FUNCTION_BLOCK EL_Template (* TEMPLATE for the rules of your equipment, EL_<Equipment>: copy it under that name, then change what says YOUR OWN, and this comment; keep the rest as it is. The logic of an equipment block: one holder at a time, outputs switched off before new ones go on, all off on release or abort, inputs reported when they change. Technical: Template: output values from its holder -> outputs (break before make); one holder at a time; all off on release or when the module aborts; inputs -> state channel when they change *)
  (* Standard: 61499-2 *)
  (* Version 0.1, 2026-09-28, Project contributors, AAU Smart Production Lab *)
  PACKAGE stoppering;
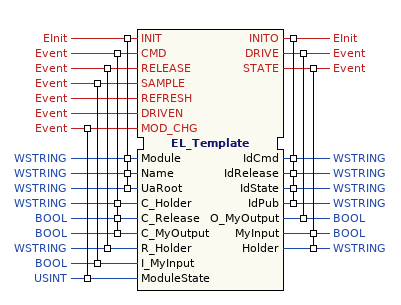
  EVENT_INPUT
    INIT : EInit WITH Module, Name, UaRoot; (* Initialise, once at start-up (the INIT chain); takes the values given with it *)
    CMD WITH C_Holder, C_Release, C_MyOutput; (* A command arrived from a holder *)
    RELEASE WITH R_Holder; (* A release arrived on the module's release channel (R_Holder) *)
    SAMPLE WITH I_MyInput; (* The inputs were read *)
    REFRESH; (* Cycle: write the outputs again *)
    DRIVEN; (* The outputs were written *)
    MOD_CHG WITH ModuleState; (* The module's state changed (its Aborting switches all off) *)
  END_EVENT
  EVENT_OUTPUT
    INITO : EInit WITH IdCmd, IdRelease, IdState, IdPub; (* Initialised: the next block of the INIT chain goes on *)
    DRIVE WITH O_MyOutput; (* Write the outputs *)
    STATE WITH MyInput, Holder; (* Publish the state (the inputs and the holder) *)
  END_EVENT
  VAR_INPUT
    Module : WSTRING; (* The module's name; its local channels are named after it (loc[<Module>/...]) *)
    Name : WSTRING; (* The equipment item's name: its local channels and OPC UA folder *)
    UaRoot : WSTRING; (* The module's OPC UA folder, e.g. /Objects/Filling *)
    C_Holder : WSTRING; (* Who sends the command *)
    C_Release : BOOL; (* Give up the equipment after this command *)
    C_MyOutput : BOOL; (* YOUR OWN, one per output pin. Commanded value of MyOutput *)
    R_Holder : WSTRING; (* Who gives up the equipment *)
    I_MyInput : BOOL; (* YOUR OWN, one per input pin. MyInput as read or received *)
    ModuleState : USINT; (* PackML state: 1 Clearing, 2 Stopped, 3 Starting, 4 Idle, 6 Execute, 7 Stopping, 8 Aborting, 9 Aborted, 15 Resetting *)
  END_VAR
  VAR_OUTPUT
    IdCmd : WSTRING; (* Local channel of the commands *)
    IdRelease : WSTRING; (* Local channel of the releases (the module's, one for all equipment) *)
    IdState : WSTRING; (* Local channel of the state *)
    IdPub : WSTRING; (* OPC UA ID of the published inputs *)
    O_MyOutput : BOOL; (* YOUR OWN, one per output pin. The value to write to MyOutput *)
    MyInput : BOOL; (* YOUR OWN, one per input pin. Template: MyInput, an input *)
    Holder : WSTRING; (* Who holds the equipment (empty: free) *)
  END_VAR
  VAR
    Publish : BOOL;
    Beat : USINT;
    LastHolder : WSTRING;
    Pending : BOOL;
    OffPending : BOOL;
    L_MyInput : BOOL; (* YOUR OWN, one per input pin *)
    N_MyOutput : BOOL; (* YOUR OWN, one per output pin *)
  END_VAR
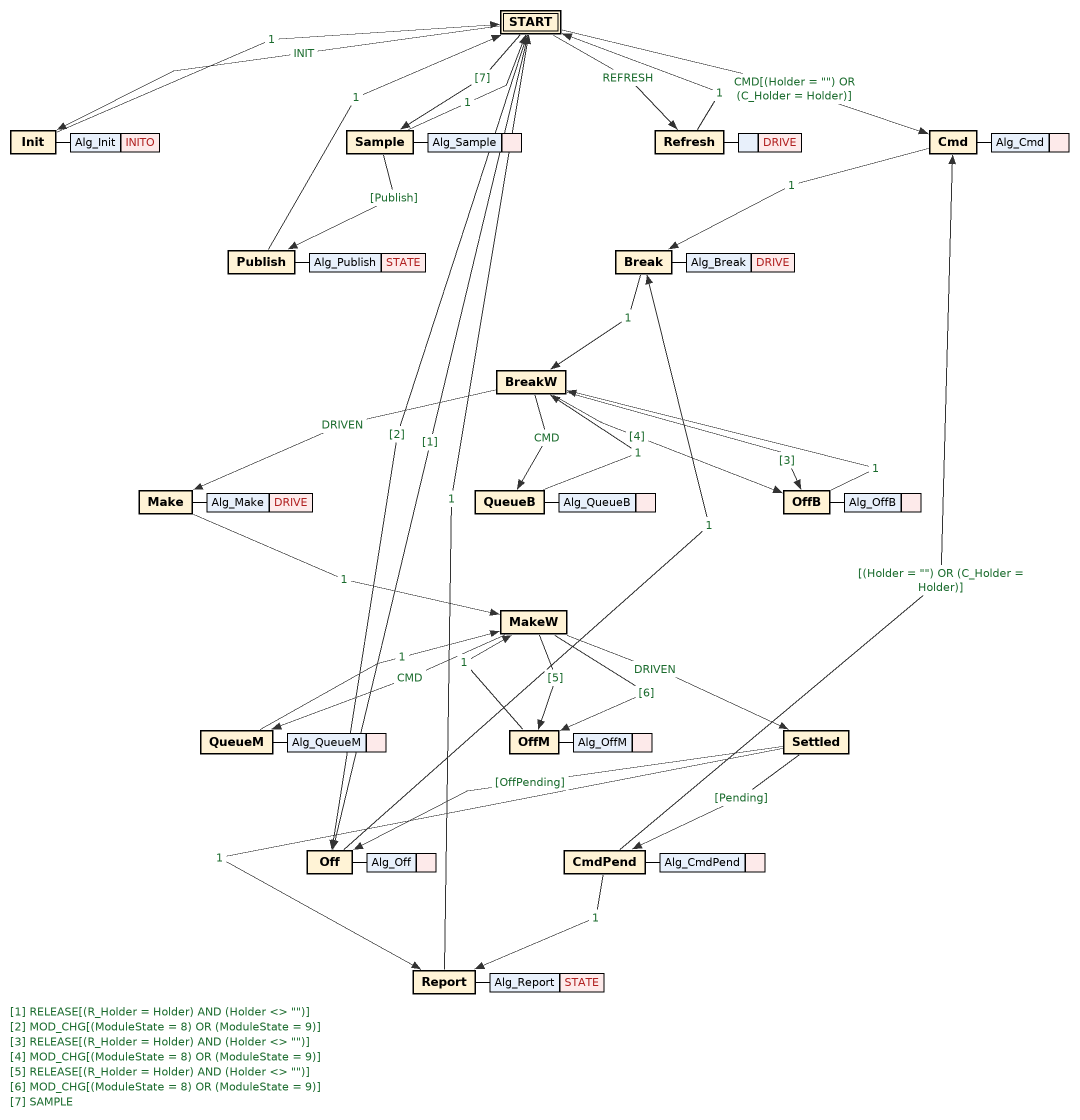
  EC_STATES
    START;
    Init : Alg_Init -> INITO;
    Sample : Alg_Sample;
    Publish : Alg_Publish -> STATE;
    Refresh : -> DRIVE;
    Cmd : Alg_Cmd;
    Off : Alg_Off;
    Break : Alg_Break -> DRIVE;
    Make : Alg_Make -> DRIVE;
    BreakW;
    MakeW;
    QueueB : Alg_QueueB;
    OffB : Alg_OffB;
    QueueM : Alg_QueueM;
    OffM : Alg_OffM;
    CmdPend : Alg_CmdPend;
    Settled;
    Report : Alg_Report -> STATE;
  END_STATES
  EC_TRANSITIONS
    START TO Init := INIT;
    START TO Sample := SAMPLE;
    START TO Refresh := REFRESH;
    START TO Cmd := CMD[(Holder = "") OR (C_Holder = Holder)];
    START TO Off := RELEASE[(R_Holder = Holder) AND (Holder <> "")];
    START TO Off := MOD_CHG[(ModuleState = 8) OR (ModuleState = 9)];
    Init TO START := 1;
    Sample TO Publish := [Publish];
    Sample TO START := 1;
    Publish TO START := 1;
    Refresh TO START := 1;
    Cmd TO Break := 1;
    Off TO Break := 1;
    Break TO BreakW := 1;
    BreakW TO Make := DRIVEN;
    Make TO MakeW := 1;
    MakeW TO Settled := DRIVEN;
    BreakW TO QueueB := CMD;
    BreakW TO OffB := RELEASE[(R_Holder = Holder) AND (Holder <> "")];
    BreakW TO OffB := MOD_CHG[(ModuleState = 8) OR (ModuleState = 9)];
    QueueB TO BreakW := 1;
    OffB TO BreakW := 1;
    MakeW TO QueueM := CMD;
    MakeW TO OffM := RELEASE[(R_Holder = Holder) AND (Holder <> "")];
    MakeW TO OffM := MOD_CHG[(ModuleState = 8) OR (ModuleState = 9)];
    QueueM TO MakeW := 1;
    OffM TO MakeW := 1;
    Settled TO Off := [OffPending];
    Settled TO CmdPend := [Pending];
    CmdPend TO Cmd := [(Holder = "") OR (C_Holder = Holder)];
    CmdPend TO Report := 1;
    Settled TO Report := 1;
    Report TO START := 1;
  END_TRANSITIONS
  ALGORITHM Alg_Init IN ST:
IdCmd := CONCAT(CONCAT(CONCAT(CONCAT("loc[", Module), "/"), Name), "/cmd]");
IdRelease := CONCAT(CONCAT("loc[", Module), "/release]");
IdState := CONCAT(CONCAT(CONCAT(CONCAT("loc[", Module), "/"), Name), "/state]");
(* YOUR OWN: the OPC UA variable of each input, with two inputs A and B: IdPub := CONCAT(CONCAT(CONCAT(CONCAT(CONCAT(CONCAT(CONCAT(CONCAT(CONCAT("opc_ua[WRITE;", UaRoot), "/Equipment/"), Name), "/A;"), UaRoot), "/Equipment/"), Name), "/B"), "]"); with none: IdPub := ""; *)
IdPub := CONCAT(CONCAT(CONCAT(CONCAT(CONCAT("opc_ua[WRITE;", UaRoot), "/Equipment/"), Name), "/MyInput"), "]");
  END_ALGORITHM
  ALGORITHM Alg_Sample IN ST:
MyInput := I_MyInput;  (* YOUR OWN: one line per input pin *)
Publish := (MyInput <> L_MyInput) OR (Holder <> LastHolder) OR (Beat >= 20);  (* YOUR OWN: one (X <> L_X) OR per input pin *)
Beat := Beat + 1;
  END_ALGORITHM
  ALGORITHM Alg_Publish IN ST:
L_MyInput := MyInput;  (* YOUR OWN: one line per input pin *)
LastHolder := Holder;
Beat := 0;
  END_ALGORITHM
  ALGORITHM Alg_Cmd IN ST:
Holder := C_Holder;
N_MyOutput := C_MyOutput;  (* YOUR OWN: one line per output pin *)
IF C_Release THEN
  Holder := "";
END_IF;
  END_ALGORITHM
  ALGORITHM Alg_Off IN ST:
N_MyOutput := FALSE;  (* YOUR OWN: one line per output pin *)
Holder := "";
OffPending := FALSE;
  END_ALGORITHM
  ALGORITHM Alg_Break IN ST:
O_MyOutput := O_MyOutput AND N_MyOutput;  (* YOUR OWN: one line per output pin *)
  END_ALGORITHM
  ALGORITHM Alg_Make IN ST:
O_MyOutput := N_MyOutput;  (* YOUR OWN: one line per output pin *)
  END_ALGORITHM
  ALGORITHM Alg_QueueB IN ST:
Pending := TRUE;
  END_ALGORITHM
  ALGORITHM Alg_OffB IN ST:
OffPending := TRUE;
  END_ALGORITHM
  ALGORITHM Alg_QueueM IN ST:
Pending := TRUE;
  END_ALGORITHM
  ALGORITHM Alg_OffM IN ST:
OffPending := TRUE;
  END_ALGORITHM
  ALGORITHM Alg_CmdPend IN ST:
Pending := FALSE;
  END_ALGORITHM
  ALGORITHM Alg_Report IN ST:
LastHolder := Holder;
Beat := 0;
  END_ALGORITHM
END_FUNCTION_BLOCK
